(*
SPDX-FileCopyrightText: © 2026 Oleksandr Tiutyk <trofimich@gmail.com>
SPDX-License-Identifier: MIT
License: https://opensource.org/license/mit
*)

(*!
<summary>Owns the lifecycle and copied diagnostic of one leaf test.</summary>
<description>
BeforeTest runs once; ExecuteTest runs according to the concrete single-cycle or multi-cycle strategy.
AfterTest runs once after normal completion, assertion failure, deadline or a caught scenario exception,
including failed preparation. Teardown must tolerate partially prepared resources. Assertions record failure
without interrupting the remaining statements of the callback. The first failure diagnostic is retained, including copied exception text/source and callback stage.
A failing exception formatter produces a stage/code fallback without replacing an earlier failure.
Exceptions from scenario hooks become one failed leaf result; catches do not roll back user side effects.
Terminal OOM propagates outside recoverable handlers and stops normal execution; teardown is not promised then.
Throwing callbacks must not use method-local resource-owning FBs that require stack unwinding.
Path-provider and reporter exceptions propagate after terminal state is committed and the stored reporter reference
is cleared. Completed callbacks are never retried.
</description>
*)

{attribute 'no_explicit_call' := 'do not call this function block directly'}
FUNCTION_BLOCK ABSTRACT TestCase EXTENDS TestElement IMPLEMENTS ITestCase
VAR
	//! <summary>Assertions bound to this case; finish one chain before starting another.</summary>
	_Assert : Assertions;	
	_Outcome : TEST_OUTCOME;
	_FailureMessage : TOF_Core.ERROR_MESSAGE;
	_Elapsed : LTIME;
	_CycleCount : UDINT;
END_VAR

(*!
<summary>Cleans up this scenario once, including after preparation or body failure.</summary>
*)
METHOD PROTECTED AfterTest
END_METHOD

(*!
<summary>Borrows the assertions bound to this running test case.</summary>
<description>Complete one immediate chain at a time; do not retain it or mutate the provider.</description>
*)
{attribute 'monitoring' := 'call'}
PROPERTY FINAL Assert : REFERENCE TO Assertions
GET
Assert REF= _Assert;
END_GET
END_PROPERTY

(*!
<summary>Prepares this scenario once per run; teardown must handle partial preparation.</summary>
*)
METHOD PROTECTED BeforeTest
END_METHOD

(*!
<summary>Counts scheduling cycles, including a deadline cycle; saturates at the UDINT maximum.</summary>
*)
{attribute 'monitoring' := 'call'}
PROPERTY FINAL CycleCount : UDINT
GET
CycleCount := _CycleCount;
END_GET
END_PROPERTY

(*!
<summary>Reports nominal time since the first scheduling cycle, initially zero.</summary>
*)
{attribute 'monitoring' := 'call'}
PROPERTY FINAL Elapsed : TIME
GET
Elapsed := TO_TIME(_Elapsed);
END_GET
END_PROPERTY

(*!
<summary>Schedules one leaf cycle and commits one result after teardown.</summary>
<description>
Scenario exceptions are converted to FAILED so the containing sequence can continue. Completion clears the
stored reporter reference before path lookup and result delivery. Exceptions from either callback propagate.
</description>
*)
// Manual stack estimate for TwinCAT. Reassess if callbacks or test workloads change.
{attribute 'estimated-stack-usage' := '16384'}
METHOD FINAL Execute
VAR
	resultReporter : ITestReporter;
	groupPath : WSTRING(255);
	exceptionCode : __SYSTEM.ExceptionCode;
	cycleResult : TEST_CYCLE_RESULT;
END_VAR
IF IsFinished THEN
	RETURN;
END_IF

IF _State = TEST_ELEMENT_STATE.READY THEN
	_State := TEST_ELEMENT_STATE.RUNNING;
	_Outcome := TEST_OUTCOME.RUNNING;
	_CycleCount := 1;
	
	_Assert.Bind(testCase := THIS^);

	__TRY
		BeforeTest();
	__CATCH(exceptionCode)
		recordRuntimeException(
			exceptionCode := exceptionCode,
			stage := 'BeforeTest',
			catchPointPOUName := __POUNAME(),
			catchPointPosition := __POSITION()
		);
	__ENDTRY

	TOF_Core.DynamicMemoryManager.RaiseIfAllocationFailed();
ELSE
	IF _CycleCount < TOF_Core.UnsignedInt32.MAX_VALUE THEN
		_CycleCount := _CycleCount + 1;
	END_IF

	_Elapsed := _Elapsed + TOF_Core.System.GetTaskCycleTime();
END_IF

_Duration := _Duration + TOF_Core.System.GetTaskCycleTime();

IF _Outcome <> TEST_OUTCOME.FAILED THEN
	__TRY
		cycleResult := RunCycle();
	__CATCH(exceptionCode)
		recordRuntimeException(
			exceptionCode := exceptionCode,
			stage := 'ExecuteTest',
			catchPointPOUName := __POUNAME(),
			catchPointPosition := __POSITION()
		);
	__ENDTRY
END_IF

TOF_Core.DynamicMemoryManager.RaiseIfAllocationFailed();

IF cycleResult <> TEST_CYCLE_RESULT.DONE AND_THEN _Outcome <> TEST_OUTCOME.FAILED THEN
	RETURN;
END_IF

__TRY
	AfterTest();
__CATCH(exceptionCode)
	recordRuntimeException(
		exceptionCode := exceptionCode,
		stage := 'AfterTest',
		catchPointPOUName := __POUNAME(),
		catchPointPosition := __POSITION()
	);
__ENDTRY

TOF_Core.DynamicMemoryManager.RaiseIfAllocationFailed();

IF _Outcome = TEST_OUTCOME.FAILED THEN
	_FailedCount := 1;
ELSE
	_Outcome := TEST_OUTCOME.PASSED;
	_PassedCount := 1;
END_IF

resultReporter := _Reporter;
_Reporter := 0;
_State := TEST_ELEMENT_STATE.COMPLETED;

IF resultReporter <> 0 THEN
	IF _Parent <> 0 THEN
		groupPath := _Parent.GetPath();
	END_IF

	resultReporter.ReportTestCaseResult(
		groupPath := groupPath,
		testName := _Name,
		outcome := _Outcome,
		duration := Duration,
		message := _FailureMessage
	);
END_IF
END_METHOD

(*!
<summary>Borrows the first copied failure diagnostic.</summary>
*)
{attribute 'monitoring' := 'call'}
PROPERTY FINAL FailureMessage : REFERENCE TO TOF_Core.ERROR_MESSAGE
GET
FailureMessage REF= _FailureMessage;
END_GET
END_PROPERTY

(*!
<summary>Reports this leaf execution outcome.</summary>
*)
{attribute 'monitoring' := 'call'}
PROPERTY FINAL Outcome : TEST_OUTCOME
GET
Outcome := _Outcome;
END_GET
END_PROPERTY

(*!
<summary>Copies the first failure while the case is running.</summary>
<description>
Does not throw for a test failure, interrupt the current callback, or change an already completed result.
</description>
*)
METHOD FINAL RecordFailure
VAR_IN_OUT CONSTANT
	message : TOF_Core.ERROR_MESSAGE;
END_VAR
IF _State <> TEST_ELEMENT_STATE.RUNNING OR_ELSE _Outcome = TEST_OUTCOME.FAILED THEN
	RETURN;
END_IF

_Outcome := TEST_OUTCOME.FAILED;
_FailureMessage := message;
END_METHOD

(*!
<summary>Copies a caught hook exception as a leaf failure without retaining its object.</summary>
<description>Preserves an earlier failure and forwards the actual catch location to diagnostic formatting.</description>
*)
METHOD PRIVATE recordRuntimeException
VAR_INPUT
	exceptionCode : __SYSTEM.ExceptionCode;
	stage : STRING;
	catchPointPOUName : STRING;
	catchPointPosition : STRING;
END_VAR
VAR
	diagnostic : TOF_Core.ERROR_MESSAGE;
END_VAR
IF _Outcome = TEST_OUTCOME.FAILED THEN
	RETURN;
END_IF

diagnostic := TestServices.FormatCaughtException(
	exceptionCode := exceptionCode,
	stage := stage,
	catchPointPOUName := catchPointPOUName,
	catchPointPosition := catchPointPosition
);
RecordFailure(message := diagnostic);
END_METHOD

(*!
<summary>Prepares fresh leaf observations without running scenario hooks.</summary>
<description>
Does not run teardown or release user resources. Call only at the lifecycle boundaries in ITestElement.
The reporter is borrowed until completion; no locks or cross-task transfer are provided.
Clears this case's outcome, diagnostic and nominal timing after common state is reset.
</description>
*)
METHOD FINAL Reset
VAR_INPUT
	reporter : ITestReporter;
END_VAR
SUPER^.Reset(reporter := reporter);

_Outcome := TEST_OUTCOME.NOT_RUN;
_FailureMessage := "";
_Elapsed := LTIME#0NS;
_CycleCount := 0;
END_METHOD

(*!
<summary>Applies the concrete scheduling strategy and returns whether the cycle finished the body.</summary>
*)
METHOD PROTECTED ABSTRACT RunCycle : TEST_CYCLE_RESULT
END_METHOD

(*!
<summary>Counts this single scenario regardless of execution state or outcome.</summary>
*)
{attribute 'monitoring' := 'call'}
PROPERTY FINAL TestCount : TOF_Core.DINT_LENGTH
GET
TestCount := 1;
END_GET
END_PROPERTY

END_FUNCTION_BLOCK

(* stored: Version 1.1.0.1
   POU TestCase: Id {a31ba67b-3136-4955-a98e-c221d790c630}, SpecialFunc None
   Folder Methods to override: Id {5136f98f-fe73-45aa-9aa8-22fc26b71a68}
   Folder Service methods: Id {a7e21a9c-64f7-4859-ad66-8eb61fb453c5}
   Method AfterTest: Id {ea6eb74d-6d37-4a53-884b-9735d2cee6ec}
   Property Assert: Id {209df581-8555-4d90-9e92-4e9dd23c4753}
   Get Get: Id {86dff3d0-5eca-434a-b68f-a96d761b4a2f}
   Method BeforeTest: Id {2155d21e-4893-47d7-a4aa-172c4bed74ea}
   Property CycleCount: Id {69d97284-2fd9-4495-807c-167c0304b62d}
   Get Get: Id {85a86a48-0389-4120-9928-ff6ad4053e71}
   Property Elapsed: Id {c3068984-8158-4fa4-ac8a-6768192d6f61}
   Get Get: Id {786808eb-177a-4daa-b8e0-a818cdcfa138}
   Method Execute: Id {5bb5d072-e228-486f-a80c-68bdefbeb2ea}
   Property FailureMessage: Id {53c0c4a4-1fd1-47f9-96b9-2c4bd55bf1c2}
   Get Get: Id {526478cc-8970-4240-a61c-23c1c29c5f99}
   Property Outcome: Id {71cd7688-473e-43fc-8a0b-ac294ef60307}
   Get Get: Id {66c3a560-7801-4af4-af5c-0868b5ecb0cf}
   Method RecordFailure: Id {a03fefe8-c08c-4d3a-b48b-b06fb20f50f9}
   Method recordRuntimeException: Id {60e6ea7f-fc70-40d6-b27c-b3fd7c82ea53}
   Method Reset: Id {7a096545-a5c2-4d84-90ff-b8fd64826a32}
   Method RunCycle: Id {c9126064-fe17-4451-994d-9a5faf603d40}
   Property TestCount: Id {06655745-6194-4112-8ff9-bf68f1de8991}
   Get Get: Id {653a1bc8-b657-4d26-8b2d-3c8b803ac45b} *)
